FUNCTION_BLOCK ASR2_SPLIT_FWD_REV (* ASR2 passthrough (Socket zu Plug) plus 2 ASR Plugs, die den Vorwaerts- und den Rueckwaerts-Kanal spiegeln *)
  (* Standard: 61499-2; Function: IN -> OUT unveraendert, zusaetzlich an FWD_OUT gespiegelt. OUT -> IN (Rueckwaerts) unveraendert, zusaetzlich an REV_OUT gespiegelt.; Description: Copyright (c) 2026 HR Agrartechnik GmbH This program and the accompanying materials are made available under the terms of the Eclipse Public License 2.0 which is available at https://www.eclipse.org/legal/epl-2.0/ SPDX-License-Identifier: EPL-2.0 *)
  (* Version 1.0, 2026-11-13, Franz Höpfinger, HR Agrartechnik GmbH, Initial Version - Luecke in der Adapter-Familie geschlossen *)
  PACKAGE adapter::events::bidirectional;
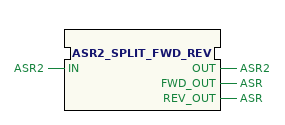
  SOCKETS
    IN : adapter::types::bidirectional::ASR2; (* bidirektionaler Eingang *)
  END_SOCKETS
  PLUGS
    OUT : adapter::types::bidirectional::ASR2; (* bidirektionaler Ausgang (Passthrough) *)
    FWD_OUT : adapter::types::unidirectional::ASR; (* spiegelt den Vorwaerts-Kanal (IN.EO* ) *)
    REV_OUT : adapter::types::unidirectional::ASR; (* spiegelt den Rueckwaerts-Kanal (OUT.EI* ) *)
  END_PLUGS
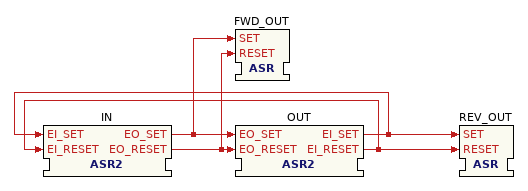
  EVENT_CONNECTIONS
    IN.EO_SET TO OUT.EO_SET;
    IN.EO_SET TO FWD_OUT.SET;
    OUT.EI_SET TO IN.EI_SET;
    OUT.EI_SET TO REV_OUT.SET;
    IN.EO_RESET TO OUT.EO_RESET;
    IN.EO_RESET TO FWD_OUT.RESET;
    OUT.EI_RESET TO IN.EI_RESET;
    OUT.EI_RESET TO REV_OUT.RESET;
  END_CONNECTIONS
END_FUNCTION_BLOCK
